(* CODESYS project cylinder.library
   DefaultNamespace: KOSTAL.AF2024.Drivers.Actuation.Cylinder
   DocFormat: reStructuredText
   Description: Handle a base cylinder device with two out and two input channels.
   Author: Frank Dümpelmann
   Title: KOSTAL.AF2024.Drivers.Actuation.Cylinder
   Version: 1.0.3.0
   Company: KOSTAL GmbH & Co.KG
   Placeholder: KOSTAL.AF2024.Drivers.Actuation.Cylinder

Project tree, tasks and I/O mapping:
  libraries: KOSTAL.AF2024.Core.functionResponse, 1.0.0.0 (KOSTAL GmbH & Co.KG); KOSTAL.AF2024.Core.ListOf, 1.0.0.0 (KOSTAL GmbH & Co.KG); KOSTAL.AF2024.Core.Process, 1.0.0.0 (KOSTAL GmbH & Co.KG); KOSTAL.AF2024.Core.Settings, 1.0.0.0 (KOSTAL GmbH & Co.KG); KOSTAL.AF2024.Core.Station, 1.0.0.0 (KOSTAL GmbH & Co.KG); KOSTAL.AF2024.Core.System, 1.0.0.0 (KOSTAL GmbH & Co.KG); KOSTAL.AF2024.Core.Text, 1.0.0.0 (KOSTAL GmbH & Co.KG); Tc2_Standard, 3.3.3.0 (Beckhoff Automation GmbH)
  Base/
    Cylinder_Base/
      function block _FB_Cylinder_Base [ST]: _fill, _mode, _moveTo_A, _moveTo_B, _pressureless, _set, conditionTime, conditionTime_ToA, conditionTime_ToB, NoLimitSwitch, sensor_A, sensor_B, valve_A, valve_B, FBmain
      interface _I_Cylinder_base: conditionTime, conditionTime_ToA, conditionTime_ToB, NoLimitSwitch, sensor_A, sensor_B, valve_A, valve_B, FBmain
      interface _I_Cylinder_base_RO: conditionTime, conditionTime_ToA, conditionTime_ToB, NoLimitSwitch, sensor_A, sensor_B, valve_A, valve_B
    Cylinder_Controlled_Base/
      function block _FB_Cylinder_Controlled_base [ST]: _manualMode_Set, _manualModeControl, _set, Error, Error_RO, errorText_overlap, errorText_timeout, ManualMode_Active, ManualMode_AutomaticRelease, ManualMode_Interlock, Name, Name_RO, overlapControl, timeout, timeoutControl, ManualMode_Reset, _fill, _moveTo_A, _moveTo_B, _pressureless, FBmain
      interface _I_Cylinder_Controlled_Base: ManualMode_Active, ManualMode_AutomaticRelease, ManualMode_Interlock, Error, Error_RO, errorText_overlap, errorText_timeout, Name, Name_RO, overlapControl, timeout, timeoutControl, ManualMode_Reset
      interface _I_Cylinder_Controlled_Base_RO: ManualMode_Active, ManualMode_AutomaticRelease, ManualMode_Interlock, Error_RO, errorText_overlap, errorText_timeout, Name_RO, overlapControl, timeout, timeoutControl
  DUT/
    Error/
      ListOf/
      interface I_T_Error: Clear, CopyFrom, active, text
      interface I_T_Error_CopyFrom: CopyFrom
      interface I_T_Error_RO: CopyTo, active, text
      function block T_Error [ST]: clear, CopyFrom, CopyTo, active, text
    Name/
      ListOf/
      interface I_T_Name: Clear, CopyFrom, device, sensor_A, sensor_B, valve_A, valve_B
      interface I_T_Name_CopyFrom: CopyFrom
      interface I_T_Name_RO: CopyTo, device, sensor_A, sensor_B, valve_A, valve_B
      function block T_Name [ST]: clear, CopyFrom, CopyTo, device, sensor_A, sensor_B, valve_A, valve_B
    StateMemory/
      ListOf/
        function block FB_ListOf_StateMemory [ST]: _get_I, _get_I_RO, _removePayLoad, _verifyMember, Add_DUT, Clear, CopyFrom, CopyTo, Delete_DUT, Find_DUT_byKey, Get_I, Get_I_RO, HasKey, Remove_DUT, MaxEntries, NumberOfMember
        interface I_ListOf_StateMemory: Add_DUT, Clear, CopyFrom, CopyTo, Delete_DUT, Get_I, Get_I_RO, NumberOfMember
        interface I_ListOf_StateMemory_CopyFrom: CopyFrom
        interface I_ListOf_StateMemory_RO: CopyTo, Get_I_RO, NumberOfMember
      interface I_T_StateMemory: Clear, CopyFrom, Key, Valve_A, Valve_B
      interface I_T_StateMemory_CopyFrom: CopyFrom
      interface I_T_StateMemory_RO: CopyTo, Key, Valve_A, Valve_B
      function block T_StateMemory [ST]: Clear, CopyFrom, CopyTo, Key, Valve_A, Valve_B
    TextHandler/
      function block FB_Text [ST]: AddVar, AddVar_UTF8, ClearVars, GetText
    data type _E_Mode
  POU/
    Cylinder/
      function block FB_Cylinder [ST]: Fill, moveTo_A, moveTo_B, Pressureless
      interface I_Cylinder: Fill, moveTo_A, moveTo_B, Pressureless
      interface I_Cylinder_RO
    Cylinder_Controlled/
      function block FB_Cylinder_Controlled [ST]: Fill, moveTo_A, moveTo_B, Pressureless
      interface I_Cylinder_Controlled: Fill, ManualMode_Reset, moveTo_A, moveTo_B, Pressureless
      interface I_Cylinder_Controlled_RO
    Cylinder_Step/
      function block FB_Cylinder_Step [ST]: FB_exit, FB_init, _addState, _StateHandling, _errorHandler, _execute, _mode, _parameterControl, ClearMemory, Fill, moveTo_A, moveTo_B, Pressureless, FBmain
      interface I_Cylinder_Step: Fill, moveTo_A, moveTo_B, Pressureless, ClearMemory
      data type ST_Manual
  Project Information/
    function F_GetCompany [ST]
    function F_GetTitle [ST]
    function F_GetVersion [ST]
  Version/
    global variables Global_Version
*)

// DUT/_E_Mode
(*
Description
===========
| Mode of cylinder control
| 0 = Normal: move to selected direction 
| 1 = Pressureless: close both valves
| 2 = Fill: open both valves  
*)
{attribute 'qualified_only'}
{attribute 'strict'}
TYPE _E_Mode :
	(
		NORMAL 			:= 0,
		PRESSURELESS	:= 1,
		FILL 			:= 2
	);
END_TYPE

// POU/Cylinder_Step/ST_Manual

TYPE ST_Manual :
STRUCT
	ManualValveMode 	: BOOL;
	ManualInterlock 	: BOOL;
	AutomaticRelease 	: BOOL;
	
	RequestManualOn		: BOOL;
	RequestManualOff	: BOOL;
	
	Valve_A				: BOOL;
	Valve_B				: BOOL;
	ResetCounter		: BYTE := 1;
	
END_STRUCT
END_TYPE

// Version/Global_Version
{attribute 'TcGenerated'}
{attribute 'no-analysis'}
{attribute 'linkalways'}
// This function has been automatically generated from the project information.
VAR_GLOBAL CONSTANT
	{attribute 'const_non_replaced'}
	stLibVersion_KOSTAL_AF2024_Drivers_Actuation_Cylinder : ST_LibVersion := (iMajor := 1, iMinor := 0, iBuild := 3, iRevision := 0, nFlags := 0, sVersion := '1.0.3.0');
END_VAR

// Base/Cylinder_Base/_FB_Cylinder_Base
{attribute 'enable_dynamic_creation'}
{attribute 'qualified_only'}
FUNCTION_BLOCK PUBLIC _FB_Cylinder_Base IMPLEMENTS _I_Cylinder_Base_RO, _I_Cylinder_Base

VAR CONSTANT
	_defTimeMin	: TIME:= TO_TIME(4294967295);	//T#0D0H0M0MS;	//define minimum default time
END_VAR

VAR
	_sensor_A	: BOOL;	//BOOL
	_sensor_B	: BOOL;	//BOOL
	_valve_A	: BOOL;	//BOOL
	_valve_B	: BOOL;	//BOOL

	_noLimitSwitch		: BOOL;
	
	_conditionTimer_moveToA	: TON;	//TON
	_conditionTime_ToA			: TIME	:= _defTimeMin;	//TIME	:= _defTimeMin - default = use common conditionTime

	_conditionTimer_moveToB	: TON;	//TON
	_conditionTime_ToB			: TIME	:= _defTimeMin;	//TIME	:= _defTimeMin - default = use common conditionTime

	_conditionTimer_moveProcess	: TON;	//TON
	_conditionTime							: TIME	:= T#100MS;	//TIME	:= T#100ms - default
	
END_VAR


METHOD PROTECTED _fill : BOOL

_fill:= FALSE;

_mode(_e_mode.FILL, FALSE, FALSE);

_conditionTimer_moveProcess.IN:= TRUE; 
_fill:= _conditionTimer_moveProcess.IN AND _conditionTimer_moveProcess.Q;
END_METHOD

METHOD PROTECTED _mode

VAR_INPUT
	mode	: _E_Mode;	//E_Mode
	to_A	: BOOL;	//BOOL
	to_B	: BOOL;	//BOOL
END_VAR
IF mode = _E_Mode.PRESSURELESS THEN

	_valve_A:= FALSE;
	_valve_B:= FALSE;

ELSIF mode = _E_Mode.FILL THEN

	_valve_A:= TRUE;
	_valve_B:= TRUE;

ELSE	//NORMAL

	_valve_A:= to_A;
	_valve_B:= to_B;
		
END_IF
END_METHOD


METHOD PROTECTED _moveTo_A : BOOL

_moveTo_A:= FALSE;

_mode(_E_Mode.NORMAL,TRUE, FALSE);

//_conditionTimer_moveToA.IN:= _sensor_A AND NOT (NOT _noSwitch AND _sensor_B);
_conditionTimer_moveToA.IN:= (_sensor_A AND NOT _sensor_B) OR _noLimitSwitch; 
 
_moveTo_A:= _conditionTimer_moveToA.IN AND _conditionTimer_moveToA.Q;
END_METHOD

METHOD PROTECTED _moveTo_B : BOOL

_moveTo_B:= FALSE;

_mode(_E_Mode.NORMAL, FALSE, TRUE);

_conditionTimer_moveToB.IN:= (_sensor_B AND NOT _sensor_A) OR _noLimitSwitch; 
_moveTo_B:= _conditionTimer_moveToB.IN AND _conditionTimer_moveToB.Q;
END_METHOD

METHOD PROTECTED _pressureless : BOOL

_pressureless:= FALSE;

_mode(_E_Mode.PRESSURELESS, FALSE, FALSE);

_conditionTimer_moveProcess.IN:= TRUE; 
_pressureless:= _conditionTimer_moveProcess.IN AND _conditionTimer_moveProcess.Q;
END_METHOD

METHOD PROTECTED _set
VAR_INPUT
END_VAR


IF _conditionTime_ToA = _defTimeMin THEN 	_conditionTimer_moveToA.PT:= _conditionTime;
ELSE																			_conditionTimer_moveToA.PT:= _conditionTime_ToA;
END_IF
_conditionTimer_moveToA();
_conditionTimer_moveToA.IN:= FALSE;	//default

IF _conditionTime_ToB = _defTimeMin THEN 	_conditionTimer_moveToB.PT:= _conditionTime;
ELSE																			_conditionTimer_moveToB.PT:= _conditionTime_ToB;
END_IF
_conditionTimer_moveToB();
_conditionTimer_moveToB.IN:= FALSE;	//default

_conditionTimer_moveProcess(IN:= , PT:= _conditionTime, Q=> , ET=> );
_conditionTimer_moveProcess.IN:= FALSE;	//default
END_METHOD

(*
Description
===========
| Minimum time before a movement function returns TRUE
*)
PROPERTY PUBLIC conditionTime : TIME
GET

conditionTime:= _conditionTime;
END_GET
SET

_conditionTime:= conditionTime;
END_SET
END_PROPERTY

(*
Description
===========
| Minimum time before a movement function returns TRUE
*)
PROPERTY PUBLIC conditionTime_ToA : TIME
GET

conditionTime_ToA:= _conditionTime_ToA;
END_GET
SET

_conditionTime_ToA:= conditionTime_ToA;
END_SET
END_PROPERTY

(*
Description
===========
| Minimum time before a movement function returns TRUE
*)
PROPERTY PUBLIC conditionTime_ToB : TIME
GET

conditionTime_ToB:= _conditionTime_ToB;
END_GET
SET

_conditionTime_ToB:= conditionTime_ToB;
END_SET
END_PROPERTY

(*
Description
===========
| TRUE: Both sensors active together result in a fault.
*)
PROPERTY PUBLIC NoLimitSwitch : BOOL
GET

NoLimitSwitch:= _noLimitSwitch;
END_GET
SET
_noLimitSwitch := NoLimitSwitch;
END_SET
END_PROPERTY

(*
Description
===========
| Sensor for home position
| Set TRUE if no sensor installed
*)
PROPERTY PUBLIC sensor_A : BOOL
GET

sensor_A:= _sensor_A;
END_GET
SET

_sensor_A:= sensor_A;
END_SET
END_PROPERTY

(*
Description
===========
| Sensor for work position
| Set TRUE if no sensor installed
*)
PROPERTY PUBLIC sensor_B : BOOL
GET

sensor_B:= _sensor_B;
END_GET
SET

_sensor_B:= sensor_B;
END_SET
END_PROPERTY

(*
Description
===========
| Valve to move cylinder to home position
*)
PROPERTY PUBLIC valve_A : BOOL
GET

valve_A:= _valve_A;
END_GET
SET

_valve_A:= valve_A;
END_SET
END_PROPERTY

(*
Description
===========
| Valve to move cylinder to work position
*)
PROPERTY PUBLIC valve_B : BOOL
GET

valve_B:= _valve_B;
END_GET
SET

_valve_B:= valve_B;
END_SET
END_PROPERTY

(*
Description
===========
| Main method, to be called cyclicly, e.g. in DeviceDefine
*)
METHOD PUBLIC FBmain
VAR_INPUT
END_VAR
	
_set();
END_METHOD

END_FUNCTION_BLOCK

// Base/Cylinder_Base/_I_Cylinder_base_RO
INTERFACE _I_Cylinder_base_RO EXTENDS KOSTAL_AF2024_Core_System.I_Interface

(*
Description
===========
| Minimum time before a movement function returns TRUE
*)
PROPERTY PUBLIC conditionTime : TIME
GET
END_GET
END_PROPERTY

(*
Description
===========
| Minimum time before a movement function returns TRUE
*)
PROPERTY PUBLIC conditionTime_ToA : TIME
GET
END_GET
END_PROPERTY

(*
Description
===========
| Minimum time before a movement function returns TRUE
*)
PROPERTY PUBLIC conditionTime_ToB : TIME
GET
END_GET
END_PROPERTY

(*
Description
===========
| TRUE: Both sensors active together result in a fault.
*)
PROPERTY PUBLIC NoLimitSwitch : BOOL
GET
END_GET
END_PROPERTY

(*
Description
===========
| Sensor for home position
| Set TRUE if no sensor installed
*)
PROPERTY PUBLIC sensor_A : BOOL
GET
END_GET
END_PROPERTY

(*
Description
===========
| Sensor for work position
| Set TRUE if no sensor installed
*)
PROPERTY PUBLIC sensor_B : BOOL
GET
END_GET
END_PROPERTY

(*
Description
===========
| Valve to move cylinder to home position
*)
PROPERTY PUBLIC valve_A : BOOL
GET
END_GET
END_PROPERTY

(*
Description
===========
| Valve to move cylinder to work position
*)
PROPERTY PUBLIC valve_B : BOOL
GET
END_GET
END_PROPERTY

END_INTERFACE

// Base/Cylinder_Base/_I_Cylinder_base
INTERFACE _I_Cylinder_base EXTENDS KOSTAL_AF2024_Core_System.I_Interface

(*
Description
===========
| Minimum time before a movement function returns TRUE
*)
PROPERTY PUBLIC conditionTime : TIME
GET
END_GET
SET
END_SET
END_PROPERTY

(*
Description
===========
| Minimum time before a movement function returns TRUE
*)
PROPERTY PUBLIC conditionTime_ToA : TIME
GET
END_GET
SET
END_SET
END_PROPERTY

(*
Description
===========
| Minimum time before a movement function returns TRUE
*)
PROPERTY PUBLIC conditionTime_ToB : TIME
GET
END_GET
SET
END_SET
END_PROPERTY

(*
Description
===========
| TRUE: Ignore Sensor inputs.
*)
PROPERTY PUBLIC NoLimitSwitch : BOOL
GET
END_GET
SET
END_SET
END_PROPERTY

(*
Description
===========
| Sensor for home position
| Set TRUE if no sensor installed
*)
PROPERTY PUBLIC sensor_A : BOOL
GET
END_GET
SET
END_SET
END_PROPERTY

(*
Description
===========
| Sensor for work position
| Set TRUE if no sensor installed
*)
PROPERTY PUBLIC sensor_B : BOOL
GET
END_GET
SET
END_SET
END_PROPERTY

(*
Description
===========
| Valve to move cylinder to home position
*)
PROPERTY PUBLIC valve_A : BOOL
GET
END_GET
SET
END_SET
END_PROPERTY

(*
Description
===========
| Valve to move cylinder to work position
*)
PROPERTY PUBLIC valve_B : BOOL
GET
END_GET
SET
END_SET
END_PROPERTY

(*
Description
===========
| Main method, to be called cyclicly, e.g. in DeviceDefine
*)
METHOD PUBLIC FBmain
VAR_INPUT
END_VAR
END_METHOD

END_INTERFACE

// Base/Cylinder_Controlled_Base/_FB_Cylinder_Controlled_base
{attribute 'enable_dynamic_creation'}
{attribute 'qualified_only'}
FUNCTION_BLOCK ABSTRACT _FB_Cylinder_Controlled_base EXTENDS _FB_Cylinder_Base IMPLEMENTS _I_Cylinder_Controlled_Base_RO, _I_Cylinder_Controlled_Base
VAR_INPUT
END_VAR
VAR_OUTPUT
END_VAR
VAR
	_timeOut			: TIME	:= T#5S;	//- default
	_timeOutTimer	: TON;
	
	_timeoutControl	: BOOL;
	_overlapControl	: BOOL;
	
	_errorText_timeout	: WSTRING;
	_errorText_overlap	: WSTRING;

	_Name		:	T_Name;
	_error	: T_Error;
	
	_textHandler	:FB_Text;
	
	//Manual control from HMI
	_automatic_A			: BOOL;
	_automatic_B			: BOOL;
	{attribute 'Cylinder_2024_V1'}
	_manual	: ST_Manual;
	
END_VAR

(*
Description
===========
| (De)activate manual valve mode
| Parameters:
| 	state : bool : TRUE = activate, FALSE = deactivate
*)
METHOD protected _manualMode_Set
VAR_INPUT
	state : bool;
END_VAR
//IF state THEN
//	_automatic_A := _valve_A;	//Store valve states before going to manual
//	_automatic_B := _valve_B;
////	_manual.ManualValveMode := TRUE;
////ELSE
////	_automatic_A 		:= FALSE;
////	_automatic_B 		:= FALSE;
////	_manual.ManualValveMode 	:= FALSE;
//END_IF
_manual.ManualValveMode := state;
END_METHOD

METHOD PROTECTED _manualModeControl
VAR_INPUT
END_VAR
IF NOT _manual.ManualValveMode THEN //Store valve states if not in manual
	_automatic_A := _valve_A;	
	_automatic_B := _valve_B;
END_IF

_manual.AutomaticRelease := (NOT (_valve_A XOR _automatic_A) AND NOT (_valve_B XOR _automatic_B));

IF _manual.RequestManualOn AND NOT _manual.ManualInterlock AND NOT _manual.ManualValveMode THEN
	//_manualMode_Set(TRUE);
	_manual.Valve_A := _valve_A;
	_manual.Valve_B := _valve_B;
	_manual.ManualValveMode := TRUE;
ELSIF _manual.RequestManualOff AND _manual.AutomaticRelease AND _manual.ManualValveMode THEN
//	_manualMode_Set(FALSE);
	_manual.ManualValveMode := FALSE;
END_IF

IF _manual.ManualValveMode AND NOT _manual.ManualInterlock THEN
	_valve_A := _manual.Valve_A;
	_valve_B := _manual.Valve_B;
END_IF
END_METHOD

METHOD PROTECTED _set
VAR_INPUT
END_VAR


SUPER^._set();


_timeOutTimer(PT:= _timeOut);
_error.active:= _timeOutTimer.Q;

_timeOutTimer.IN:= FALSE;	//default

_error.clear();
END_METHOD

(*
Description
===========
| See documentation of FB_error
| **Attention:** Errors are reset in FB_Main. Check errors before FB_Main is called!
*)
PROPERTY PUBLIC Error : I_T_Error
GET

Error := _error;
END_GET
END_PROPERTY

PROPERTY PUBLIC Error_RO : I_T_Error_RO
GET

Error_RO:= _error;
END_GET
END_PROPERTY

(*
Description
===========
| Message Text for overlap error
*)
PROPERTY PUBLIC errorText_overlap : KOSTAL_AF2024_Core_Settings.T_MaxString
GET

errorText_overlap:= _errorText_overlap;
END_GET
SET

_errorText_overlap:= errorText_overlap;
END_SET
END_PROPERTY

(*
Description
===========
| Message Text for timeout error
*)
PROPERTY PUBLIC errorText_timeout : KOSTAL_AF2024_Core_Settings.T_MaxString
GET

errorText_Timeout:= _errorText_timeout;
END_GET
SET

_errorText_Timeout:= errorText_timeout;
END_SET
END_PROPERTY

(*
Description
===========
| TRUE if manual control is activated for this cylinder
*)
PROPERTY PUBLIC ManualMode_Active : BOOL
GET
ManualMode_Active := _manual.ManualValveMode;
END_GET
END_PROPERTY

(*
Description
===========
| True if manual valve state equals automatic valve state
| -> Enable automatic mode 
*)
// 
PROPERTY PUBLIC ManualMode_AutomaticRelease : BOOL
GET
ManualMode_AutomaticRelease := _manual.AutomaticRelease;
END_GET
END_PROPERTY

(*
Description
===========
| Interlock manual cylinder control
*)
PROPERTY PUBLIC ManualMode_Interlock : BOOL
GET
ManualMode_Interlock := _manual.ManualInterlock;
END_GET
SET
_manual.ManualInterlock := ManualMode_Interlock;
END_SET
END_PROPERTY

PROPERTY PUBLIC Name : I_T_Name
GET

Name:= _Name;
END_GET
END_PROPERTY

(*
Description
===========
| Naming of cilinders and componets (see documentation of FB_name)
*)
PROPERTY PUBLIC Name_RO : I_T_Name_RO
GET

Name_RO := _Name;
END_GET
END_PROPERTY

(*
Description
===========
| TRUE: Both sensors active together result in a fault.
*)
PROPERTY PUBLIC overlapControl : BOOL
GET

overlapControl:= _overlapControl;
END_GET
SET

_overlapControl:= overlapControl;
END_SET
END_PROPERTY

(*
Description
===========
| Time for timeoutControl
| Default: 5s
*)
PROPERTY PUBLIC timeout : TIME
GET

timeout:= _timeOut;
END_GET
SET

_timeout:= timeOut;
END_SET
END_PROPERTY

(*
Description
===========
| TRUE: generate error when movement is not finished after a certain time
*)
PROPERTY PUBLIC timeoutControl : BOOL
GET

timeoutControl:= _timeoutControl;
END_GET
SET

_timeoutControl:= timeoutControl;
END_SET
END_PROPERTY

METHOD Public ManualMode_Reset : BOOL
VAR_INPUT
END_VAR

_manualMode_Set(FALSE);
_manual.Valve_A := _manual.Valve_B := FALSE;
_manual.ResetCounter := LIMIT(1, _manual.ResetCounter + 1, 254);

ManualMode_Reset := THIS^._pressureless();
END_METHOD

METHOD PROTECTED _fill : BOOL

_fill:= SUPER^._fill();

_timeOutTimer(IN:= NOT _conditionTimer_moveProcess.IN AND _timeoutControl, PT:= _timeOut);

IF _overlapControl AND _sensor_A AND _sensor_B AND NOT _noLimitSwitch THEN

	_error.active:= TRUE;

	_textHandler.clearVars();
	_textHandler.AddVar(Name_RO.sensor_A);
	_textHandler.AddVar(Name_RO.sensor_B);
	_error.text:=  _textHandler.getText(errorText_overlap);

ELSE

	_error.active:= FALSE;
	_error.text:= "";
	
END_IF
END_METHOD

METHOD PROTECTED _moveTo_A : BOOL

_moveTo_A:= SUPER^._moveTo_A();


_timeOutTimer(IN:= NOT _conditionTimer_moveToA.IN AND _timeoutControl, PT:= _timeOut);

IF _overlapControl AND _sensor_A AND _sensor_B AND NOT _noLimitSwitch THEN

	_error.active:= TRUE;
	
	_textHandler.clearVars();
	_textHandler.AddVar(Name_RO.sensor_A);
	_textHandler.AddVar(Name_RO.sensor_B);
	_error.text:=  _textHandler.GetText(errorText_overlap);

ELSIF _timeOutTimer.Q THEN

	_error.active:= TRUE;

	_textHandler.clearVars();
	_textHandler.AddVar(Name_RO.sensor_A);
	_error.text:=  _textHandler.GetText(errorText_timeout);

ELSE

	_error.active:= FALSE;
	_error.text:= "";
	
END_IF
END_METHOD

METHOD PROTECTED _moveTo_B : BOOL

_moveTo_B:= SUPER^._moveTo_B();


_timeOutTimer(IN:= NOT _conditionTimer_moveToB.IN AND _timeoutControl, PT:= _timeOut);

IF _overlapControl AND _sensor_A AND _sensor_B AND NOT _noLimitSwitch THEN

	_error.active:= TRUE;

	_textHandler.clearVars();
	_textHandler.AddVar(Name_RO.sensor_A);
	_textHandler.AddVar(Name_RO.sensor_B);
	_error.text:=  _textHandler.getText(errorText_overlap);

ELSIF _timeOutTimer.Q THEN

	_error.active:= TRUE;

	_textHandler.clearVars();
	_textHandler.AddVar(Name_RO.sensor_B);
	_error.text:=  _textHandler.getText(errorText_timeout);

ELSE

	_error.active:= FALSE;
	_error.text:= "";
	
END_IF
END_METHOD

METHOD PROTECTED _pressureless : BOOL

_pressureless:= SUPER^._pressureless();

_timeOutTimer(IN:= NOT _conditionTimer_moveProcess.IN AND _timeoutControl, PT:= _timeOut);

IF _overlapControl AND _sensor_A AND _sensor_B AND NOT _noLimitSwitch THEN

	_error.active:= TRUE;

	_textHandler.clearVars();
	_textHandler.AddVar(Name_RO.sensor_A);
	_textHandler.AddVar(Name_RO.sensor_B);
	_error.text:=  _textHandler.getText(errorText_overlap);

ELSE

	_error.active:= FALSE;
	_error.text:= "";
	
END_IF
END_METHOD

(*
Description
===========
| Main method, to be called cyclicly, e.g. in DeviceDefine
*)
METHOD PUBLIC FBmain
VAR_INPUT
END_VAR
SUPER^.FBmain();
_manualModeControl();
END_METHOD

END_FUNCTION_BLOCK

// Base/Cylinder_Controlled_Base/_I_Cylinder_Controlled_Base_RO
INTERFACE _I_Cylinder_Controlled_Base_RO EXTENDS _I_Cylinder_Base_RO

PROPERTY PUBLIC ManualMode_Active : BOOL
GET
END_GET
END_PROPERTY

//Manual valve state = automatic valve state -> Release automatic mode
PROPERTY PUBLIC ManualMode_AutomaticRelease : BOOL
GET
END_GET
END_PROPERTY

PROPERTY PUBLIC ManualMode_Interlock : BOOL
GET
END_GET
END_PROPERTY

PROPERTY PUBLIC Error_RO : I_T_Error_RO
GET
END_GET
END_PROPERTY

(*
Description
===========
| Message Text for overlap error
*)
PROPERTY PUBLIC errorText_overlap : KOSTAL_AF2024_Core_Settings.T_MaxString
GET
END_GET
SET
END_SET
END_PROPERTY

(*
Description
===========
| Message Text for timeout error
*)
PROPERTY PUBLIC errorText_timeout : KOSTAL_AF2024_Core_Settings.T_MaxString
GET
END_GET
END_PROPERTY

(*
Description
===========
| Naming of cilinders and componets (see documentation of FB_name)
*)
{attribute 'obsolete' := 'use instead property IName or method LinkName()!'} 
PROPERTY PUBLIC Name_RO : I_T_Name_RO
GET
END_GET
END_PROPERTY

(*
Description
===========
| TRUE: Both sensors active together result in a fault.
*)
PROPERTY PUBLIC overlapControl : BOOL
GET
END_GET
END_PROPERTY

(*
Description
===========
| Time for timeoutControl
| Default: 5s
*)
PROPERTY PUBLIC timeout : TIME
GET
END_GET
END_PROPERTY

(*
Description
===========
| TRUE: generate error when movement is not finished after a certain time
*)
PROPERTY PUBLIC timeoutControl : BOOL
GET
END_GET
END_PROPERTY

END_INTERFACE

// DUT/Error/I_T_Error_RO
(*
	Read only Interface from DUT
*)
INTERFACE I_T_Error_RO  EXTENDS KOSTAL_AF2024_Core_System.I_Interface

METHOD PUBLIC CopyTo
VAR_INPUT
	IN	: I_T_Error_CopyFrom;
END_VAR
END_METHOD

(*
Description
===========
| Error is active
*)
PROPERTY PUBLIC active : BOOL
GET
END_GET
END_PROPERTY

(*
Description
===========
| Text of error message
*)
PROPERTY PUBLIC text : KOSTAL_AF2024_Core_Settings.T_MaxString
GET
END_GET
END_PROPERTY

END_INTERFACE

// DUT/Error/I_T_Error_CopyFrom
INTERFACE I_T_Error_CopyFrom EXTENDS KOSTAL_AF2024_Core_System.I_Interface

METHOD PUBLIC CopyFrom
VAR_INPUT
	IN	: I_T_Error_RO;
END_VAR
END_METHOD

END_INTERFACE

// DUT/Name/I_T_Name_RO
(*
	Read only Interface from DUT
*)
INTERFACE I_T_Name_RO  EXTENDS KOSTAL_AF2024_Core_System.I_Interface

METHOD PUBLIC CopyTo
VAR_INPUT
	IN	: I_T_Name_CopyFrom;
END_VAR
END_METHOD

(*
Description
===========
| Name of the cylinder
*)
PROPERTY PUBLIC device : KOSTAL_AF2024_Core_Settings.T_MaxString
GET
END_GET
END_PROPERTY

(*
Description
===========
| Name of the cylinder's home position sensor
*)
PROPERTY PUBLIC sensor_A : KOSTAL_AF2024_Core_Settings.T_MaxString
GET
END_GET
END_PROPERTY

(*
Description
===========
| Name of the cylinder's work position sensor
*)
PROPERTY PUBLIC sensor_B : KOSTAL_AF2024_Core_Settings.T_MaxString
GET
END_GET
END_PROPERTY

(*
Description
===========
| Name of the cylinder's home position actuator
*)
PROPERTY PUBLIC valve_A : KOSTAL_AF2024_Core_Settings.T_MaxString
GET
END_GET
END_PROPERTY

(*
Description
===========
| Name of the cylinder's work position actuator
*)
PROPERTY PUBLIC valve_B : KOSTAL_AF2024_Core_Settings.T_MaxString
GET
END_GET
END_PROPERTY

END_INTERFACE

// DUT/Name/I_T_Name_CopyFrom
INTERFACE I_T_Name_CopyFrom EXTENDS KOSTAL_AF2024_Core_System.I_Interface

METHOD PUBLIC CopyFrom
VAR_INPUT
	IN	: I_T_Name_RO;
END_VAR
END_METHOD

END_INTERFACE

// Base/Cylinder_Controlled_Base/_I_Cylinder_Controlled_Base
INTERFACE _I_Cylinder_Controlled_Base EXTENDS _I_Cylinder_base

PROPERTY PUBLIC ManualMode_Active : BOOL
GET
END_GET
END_PROPERTY

//Manual valve state = automatic valve state -> Release automatic mode
PROPERTY PUBLIC ManualMode_AutomaticRelease : BOOL
GET
END_GET
END_PROPERTY

PROPERTY PUBLIC ManualMode_Interlock : BOOL
GET
END_GET
SET
END_SET
END_PROPERTY

(*
Description
===========
| See documentation of FB_error
| **Attention:** Errors are reset in FB_Main. Check errors before FB_Main is called!
*)
PROPERTY PUBLIC Error : I_T_Error
GET
END_GET
END_PROPERTY

PROPERTY PUBLIC Error_RO : I_T_Error_RO
GET
END_GET
END_PROPERTY

(*
Description
===========
| Message Text for overlap error
*)
PROPERTY PUBLIC errorText_overlap : KOSTAL_AF2024_Core_Settings.T_MaxString
GET
END_GET
SET
END_SET
END_PROPERTY

(*
Description
===========
| Message Text for timeout error
*)
PROPERTY PUBLIC errorText_timeout : KOSTAL_AF2024_Core_Settings.T_MaxString
GET
END_GET
SET
END_SET
END_PROPERTY

PROPERTY PUBLIC Name : I_T_Name
GET
END_GET
END_PROPERTY

(*
Description
===========
| Naming of cilinders and componets (see documentation of FB_name)
*)
{attribute 'obsolete' := 'use instead property IName or method LinkName()!'} 
PROPERTY PUBLIC Name_RO : I_T_Name_RO
GET
END_GET
END_PROPERTY

(*
Description
===========
| TRUE: Both sensors active together result in a fault.
*)
PROPERTY PUBLIC overlapControl : BOOL
GET
END_GET
SET
END_SET
END_PROPERTY

(*
Description
===========
| Time for timeoutControl
| Default: 5s
*)
PROPERTY PUBLIC timeout : TIME
GET
END_GET
SET
END_SET
END_PROPERTY

(*
Description
===========
| TRUE: generate error when movement is not finished after a certain time
*)
PROPERTY PUBLIC timeoutControl : BOOL
GET
END_GET
SET
END_SET
END_PROPERTY

METHOD Public ManualMode_Reset : BOOL
VAR_INPUT
END_VAR
END_METHOD

END_INTERFACE

// DUT/Error/I_T_Error
(*
	Full qualified access Interface from DUT
*)
INTERFACE I_T_Error EXTENDS I_T_Error_RO

METHOD PUBLIC Clear
END_METHOD

METHOD PUBLIC CopyFrom
VAR_INPUT
	IN	: I_T_Error_RO;
END_VAR
END_METHOD

(*
Description
===========
| Error is active
*)
PROPERTY PUBLIC active : BOOL
SET
END_SET
END_PROPERTY

(*
Description
===========
| Text of error message
*)
PROPERTY PUBLIC text : KOSTAL_AF2024_Core_Settings.T_MaxString
SET
END_SET
END_PROPERTY

END_INTERFACE

// DUT/Name/I_T_Name
(*
	Full qualified access Interface from DUT
*)
INTERFACE I_T_Name EXTENDS I_T_Name_RO

METHOD PUBLIC Clear : BOOL
VAR_INPUT
END_VAR
END_METHOD

METHOD PUBLIC CopyFrom
VAR_INPUT
	IN	: I_T_Name_RO;
END_VAR
END_METHOD

(*
Description
===========
| Name of the cylinder
*)
PROPERTY PUBLIC device : KOSTAL_AF2024_Core_Settings.T_MaxString
SET
END_SET
END_PROPERTY

(*
Description
===========
| Name of the cylinder's home position sensor
*)
PROPERTY PUBLIC sensor_A : KOSTAL_AF2024_Core_Settings.T_MaxString
SET
END_SET
END_PROPERTY

(*
Description
===========
| Name of the cylinder's work position sensor
*)
PROPERTY PUBLIC sensor_B : KOSTAL_AF2024_Core_Settings.T_MaxString
SET
END_SET
END_PROPERTY

(*
Description
===========
| Name of the cylinder's home position actuator
*)
PROPERTY PUBLIC valve_A : KOSTAL_AF2024_Core_Settings.T_MaxString
SET
END_SET
END_PROPERTY

(*
Description
===========
| Name of the cylinder's work position actuator
*)
PROPERTY PUBLIC valve_B : KOSTAL_AF2024_Core_Settings.T_MaxString
SET
END_SET
END_PROPERTY

END_INTERFACE

// DUT/Name/T_Name
(*

:Author: Frank Dümpelmann <f.duempelmann@kostal.com>, Martin Hundt <m.hundt@kostal.com>
:Date: 2018-11-19

Function
========
| Data type for naming cylinders and their components (valves, sensors)

Methods and Properties
======================
| See bottom of this document for a detailed description of each method or property
*)

{attribute 'enable_dynamic_creation'}
{attribute 'qualified_only'}
FUNCTION_BLOCK T_Name IMPLEMENTS I_T_Name_RO, I_T_Name, I_T_Name_CopyFrom

VAR
	_device		: KOSTAL_AF2024_Core_Settings.T_MaxString;
	_sensor_A	: KOSTAL_AF2024_Core_Settings.T_MaxString;
	_sensor_B	: KOSTAL_AF2024_Core_Settings.T_MaxString;
	_valve_A	: KOSTAL_AF2024_Core_Settings.T_MaxString;
	_valve_B	: KOSTAL_AF2024_Core_Settings.T_MaxString;
END_VAR

(*
Description
===========
| Clear all naming
*)
METHOD clear : BOOL
VAR_INPUT
END_VAR

_device		:= "";
_sensor_A	:= "";
_sensor_B	:= "";
_valve_A	:= "";
_valve_B	:= "";
END_METHOD

METHOD PUBLIC CopyFrom
VAR_INPUT
	IN	: I_T_Name_RO;
END_VAR

IF IN = 0 THEN RETURN;	END_IF

_device		:= IN.device;
_sensor_A	:= IN.sensor_A;
_sensor_B	:= IN.sensor_B;
_valve_A	:= IN.valve_A;
_valve_B	:= IN.valve_B;
END_METHOD

METHOD PUBLIC CopyTo
VAR_INPUT
	IN	: I_T_Name_CopyFrom;
END_VAR

IF IN = 0 THEN RETURN;	END_IF

IN.CopyFrom(THIS^);
END_METHOD

(*
Description
===========
| Name of the cylinder
*)
PROPERTY PUBLIC device : KOSTAL_AF2024_Core_Settings.T_MaxString
GET

device:= _device;
END_GET
SET

_device:= device;
END_SET
END_PROPERTY

(*
Description
===========
| Name of the cylinder's home position sensor
*)
PROPERTY PUBLIC sensor_A : KOSTAL_AF2024_Core_Settings.T_MaxString
GET

sensor_A:= _sensor_A;
END_GET
SET

_sensor_A:= sensor_A;
END_SET
END_PROPERTY

(*
Description
===========
| Name of the cylinder's work position sensor
*)
PROPERTY PUBLIC sensor_B : KOSTAL_AF2024_Core_Settings.T_MaxString
GET

sensor_B:= _sensor_B;
END_GET
SET

_sensor_B:= sensor_B;
END_SET
END_PROPERTY

(*
Description
===========
| Name of the cylinder's home position actuator
*)
PROPERTY PUBLIC valve_A : KOSTAL_AF2024_Core_Settings.T_MaxString
GET

valve_A:= _valve_A;
END_GET
SET

_valve_A:= valve_A;
END_SET
END_PROPERTY

(*
Description
===========
| Name of the cylinder's work position actuator
*)
PROPERTY PUBLIC valve_B : KOSTAL_AF2024_Core_Settings.T_MaxString
GET

valve_B:= _valve_B;
END_GET
SET

_valve_B:= valve_B;
END_SET
END_PROPERTY

END_FUNCTION_BLOCK

// DUT/Error/T_Error
(*

:Author: Frank Dümpelmann <f.duempelmann@kostal.com>, Martin Hundt <m.hundt@kostal.com>
:Date: 2018-11-19

Function
========
| Data type for error messages

Methods and Properties
======================
| See bottom of this document for a detailed description of each method or property
*)
{attribute 'enable_dynamic_creation'}
{attribute 'qualified_only'}
FUNCTION_BLOCK T_Error IMPLEMENTS I_T_Error_RO, I_T_Error, I_T_Error_CopyFrom

VAR
	_active	: BOOL;
	_text		: KOSTAL_AF2024_Core_Settings.T_MaxString;
END_VAR

METHOD PUBLIC Clear

_active	:= FALSE;
_text		:= "";
END_METHOD

METHOD PUBLIC CopyFrom
VAR_INPUT
	IN	: I_T_Error_RO;
END_VAR

IF IN = 0 THEN RETURN;	END_IF

_active	:= IN.active;
_text		:= IN.text;
END_METHOD

METHOD PUBLIC CopyTo
VAR_INPUT
	IN	: I_T_Error_CopyFrom;
END_VAR

IF IN = 0 THEN RETURN;	END_IF

IN.CopyFrom(THIS^);
END_METHOD

(*
Description
===========
| Error is active
*)
PROPERTY PUBLIC active : BOOL
GET

active:= _active;
END_GET
SET

_active:= active;
END_SET
END_PROPERTY

(*
Description
===========
| Text of error message
*)
PROPERTY PUBLIC text : KOSTAL_AF2024_Core_Settings.T_MaxString
GET

text:= _text;
END_GET
SET

_text:= text;
END_SET
END_PROPERTY

END_FUNCTION_BLOCK

// DUT/TextHandler/FB_Text
FUNCTION_BLOCK INTERNAL FB_Text EXTENDS Kostal_AF2024_Core_Text._FB_Base
VAR_INPUT
END_VAR
VAR_OUTPUT
END_VAR
VAR
END_VAR

METHOD AddVar : BOOL
VAR_INPUT
	Text	: KOSTAL_AF2024_Core_Settings.T_MaxString;
END_VAR

AddVar:= _Variables.addLine(Text);
END_METHOD

METHOD AddVar_UTF8 : BOOL
VAR_INPUT
	Text	: KOSTAL_AF2024_Core_Settings.T_MaxString;
END_VAR



AddVar_UTF8:= _Variables.addLine(Text);
END_METHOD

METHOD ClearVars

_Variables.clear();
END_METHOD

METHOD GetText : KOSTAL_AF2024_Core_Settings.T_MaxString

VAR_INPUT
	Text	: KOSTAL_AF2024_Core_Settings.T_MaxString;
END_VAR

GetText:= "";

IF Text = "" THEN RETURN;	END_IF

GetText:= _combine(Text);
END_METHOD

END_FUNCTION_BLOCK

// DUT/StateMemory/ListOf/FB_ListOf_StateMemory
(*
	A template for creating a list of typed classes (FBs)
*)
FUNCTION_BLOCK FB_ListOf_StateMemory EXTENDS KOSTAL_AF2024_Core_ListOf._FB_Object_Base  IMPLEMENTS I_ListOf_StateMemory_RO, I_ListOf_StateMemory_CopyFrom, I_ListOf_StateMemory

VAR
	//Use the {_Dummy} to ensure that a valid interface is always returned.
	_Dummy			: T_StateMemory;
	_MaxEntries	: UDINT:= UDINT#128;
END_VAR

(*
	Returns the typed owner interface in the reference variable.
	In the event of an error, the return value becomes FALSE and the interface refers to the {_Dummy}.
*)
METHOD PROTECTED _get_I : BOOL

VAR_INPUT
	Member		: KOSTAL_AF2024_Core_System.I_Interface;
	rFound_I	: REFERENCE TO I_T_StateMemory;
	rResult		: KOSTAL_AF2024_Core_functionResponse.I_T_functionResponse_Owner;
END_VAR

VAR
	_iObj			: I_T_StateMemory;
	_Success	: BOOL;
END_VAR

IF NOT SUPER^._verifyMember(Member, rResult)	THEN 
	IF __ISVALIDREF(rFound_I)	THEN	rFound_I:= _Dummy;	END_IF
	RETURN;	
END_IF

_Success:= __QUERYINTERFACE(Member, _iObj);

//return dummy if no valid DUT is found
IF NOT _Success OR (_iObj = 0)	THEN	

	IF __ISVALIDREF(rFound_I)	THEN	rFound_I:= _Dummy;	END_IF	
	IF rResult <> 0						THEN	rResult.success:= FALSE;	
																	rResult.status:= "__QueryInterface failed - return Dummy";	
	END_IF	

	RETURN;	

END_IF

IF __ISVALIDREF(rFound_I)	THEN	rFound_I:= _iObj;	END_IF
IF rResult <> 0						THEN	rResult.success:= TRUE;
																rResult.status:= "Successful";
END_IF

_get_I:= TRUE;
END_METHOD

(*
	Returns the typed interface in the reference variable.
	In the event of an error, the return value becomes FALSE and the interface refers to the {_Dummy}.
*)
METHOD PROTECTED _get_I_RO : BOOL

VAR_INPUT
	Member		: KOSTAL_AF2024_Core_System.I_Interface;
	rFound_I	: REFERENCE TO I_T_StateMemory_RO;
	rResult		: KOSTAL_AF2024_Core_functionResponse.I_T_functionResponse_Owner;
END_VAR

VAR
	_iObj	: I_T_StateMemory_RO;
	_Success: BOOL;
END_VAR

IF NOT SUPER^._verifyMember(Member, rResult)	THEN 
	IF __ISVALIDREF(rFound_I)	THEN	rFound_I:= _Dummy;	END_IF
	RETURN;	
END_IF

_Success:= __QUERYINTERFACE(Member, _iObj);

//return dummy if no valid DUT is found
IF NOT _Success OR (_iObj = 0)	THEN	

	IF __ISVALIDREF(rFound_I)	THEN	rFound_I:= _Dummy;	END_IF	
	IF rResult <> 0						THEN	rResult.success:= FALSE;		
																	rResult.status:= "__QueryInterface failed - return Dummy";	
	END_IF	

	RETURN;	

END_IF

IF __ISVALIDREF(rFound_I)	THEN	rFound_I:= _iObj;	END_IF
IF rResult <> 0						THEN	rResult.success:= TRUE;
																rResult.status:= "Successful";
END_IF

_get_I_RO:= TRUE;
END_METHOD

(*
	Cleans the custom class {FB_DUT} and removes it from memory.
*)
METHOD PROTECTED  _removePayLoad : BOOL
VAR_INPUT
	Member	: KOSTAL_AF2024_Core_System.I_Interface;
	Result	: KOSTAL_AF2024_Core_functionResponse.I_T_functionResponse_Owner;
END_VAR

VAR
	_iObj			: I_T_StateMemory;
	_pFB_DUT	:	POINTER TO T_StateMemory;
	_Success	: BOOL;
END_VAR


IF NOT SUPER^._removePayload(Member, Result)	THEN RETURN;	END_IF

_Success:= __QUERYINTERFACE(Member, _iObj);

IF NOT _Success	THEN	RETURN;	END_IF
IF _iObj = 0		THEN	RETURN;	END_IF

_iObj.Clear();

_Success  := __QUERYPOINTER(_iObj, _pFB_DUT);

IF NOT _Success	THEN	RETURN;	END_IF
IF _pFB_DUT = 0	THEN	RETURN;	END_IF

__DELETE(_pFB_DUT);
END_METHOD

(*
	Overload the method from the base class to verify the custom interface. 
	The local method {_get_I_Owner()} is used for this.
*)
METHOD PROTECTED _verifyMember : BOOL
VAR_INPUT
	Member	: KOSTAL_AF2024_Core_System.I_Interface;
	Result	: KOSTAL_AF2024_Core_functionResponse.I_T_functionResponse_Owner;
END_VAR


_verifyMember:= _get_I(Member, 0, Result);
END_METHOD

(*
	Add a new instance of FB_Dut and copy content from [IN] to the new instance
*)
METHOD PUBLIC Add_DUT : BOOL
VAR_INPUT
	IN				: I_T_StateMemory_RO;
	Response	: KOSTAL_AF2024_Core_functionResponse.I_T_functionResponse_Owner;
END_VAR

VAR
	_iDUT	: I_T_StateMemory;
	_pDUT: POINTER TO T_StateMemory;
	_response: KOSTAL_AF2024_Core_functionResponse.T_functionResponse;
	_udi: UDINT;
END_VAR

_response.clear();

IF IN = 0 THEN
	IF Response <> 0 THEN	Response.success:= FALSE;	Response.status:= "IN Parameter is invalid";	END_IF
	RETURN;
END_IF

IF _Count	> _MaxEntries THEN 
	IF Response <> 0 THEN	Response.success:= FALSE;	Response.status:= "Max entries overflow";	END_IF
	RETURN;	
END_IF

_pDUT:= __NEW(T_StateMemory);

IF _pDUT = 0 THEN
	_response.status:= "cannot create new object";
	IF Response <> 0 THEN	Response.CopyFrom(_response);	END_IF
	RETURN;
END_IF

_pDUT^.CopyFrom(IN);

SUPER^._addMember(_pDUT^, _response);

IF Response <> 0 THEN	Response.CopyFrom(_response);	END_IF

Add_DUT:= _response.success;
END_METHOD

(*
	Makes the protected method public.
*)
METHOD Clear

SUPER^._clear();
END_METHOD

(*
	Copies the contents of another list {IN} into its own memory.
*)
METHOD PUBLIC CopyFrom
VAR_INPUT
	IN	: I_ListOf_StateMemory_RO;
END_VAR

VAR
	_udi	: UDINT;
	_IDUT	: I_T_StateMemory_RO;
END_VAR
IF IN = 0 THEN RETURN;	END_IF

_clear();

FOR _udi:= 1 TO IN.NumberOfMember DO
	IF IN.Get_I_RO(_udi, _IDUT, 0)	THEN	Add_DUT(_IDUT, 0);	END_IF
END_FOR
END_METHOD

(*
	Copies the own content into another list created at the parameter {IN}.
*)
METHOD PUBLIC CopyTo
VAR_INPUT
	IN	: I_ListOf_StateMemory_CopyFrom;
END_VAR

IF IN = 0 THEN RETURN;	END_IF

IN.CopyFrom(THIS^);
END_METHOD

(*
	Deletes the class specified with the {Number} from the list.
*)
METHOD PUBLIC Delete_DUT : BOOL
VAR_INPUT
	Number		: UDINT;	//Number of DUT in List
	Response	: KOSTAL_AF2024_Core_functionResponse.I_T_functionResponse_Owner;
END_VAR

VAR
	_response	: KOSTAL_AF2024_Core_functionResponse.T_functionResponse;
	_Success	: BOOL;
	_Member		: KOSTAL_AF2024_Core_System.I_Interface;
END_VAR

IF Number = 0 THEN
	_response.clear(); _response.status:= "Number is out of range (1..n)"; 
	IF Response <> 0 THEN	Response.CopyFrom(_response);	END_IF
	RETURN;
END_IF

Delete_DUT:= SUPER^._removeMemberByIndex(Number - 1, _response);

IF Response <> 0 THEN	Response.CopyFrom(_response);	END_IF

Delete_DUT:= _response.success;
END_METHOD

METHOD Find_DUT_byKey : BOOL
VAR_INPUT
	Key	: ULINT;
	rFound_I	: REFERENCE TO I_T_StateMemory_RO;
END_VAR

VAR
	_udi: UDINT;
	_iMem				: KOSTAL_AF2024_Core_System.I_Interface;
	_iStateMem	: I_T_StateMemory_RO;
	_Success: BOOL;
END_VAR

IF _Count = 0 THEN	rFound_I:= _Dummy;	Find_DUT_byKey:= FALSE;	RETURN;	END_IF

FOR _udi:= _Count - 1 TO 0 BY -1 DO 

	IF _findMemberByIndex(_udi, _iMem, 0) AND_THEN _iMem <> 0 THEN 

		_Success:= __QUERYINTERFACE(_iMem, _iStateMem);
		
		//return dummy if no valid DUT is found
		IF NOT _Success OR_ELSE (_iStateMem = 0)	THEN	
		
			IF __ISVALIDREF(rFound_I)	THEN	rFound_I:= _Dummy;	Find_DUT_byKey:= FALSE; END_IF	
			RETURN;	

		ELSE

			IF _iStateMem.Key = Key THEN
					
				IF __ISVALIDREF(rFound_I) THEN	rFound_I:= _iStateMem;	Find_DUT_byKey:= TRUE;	RETURN;	END_IF
		
			END_IF


		END_IF
	
	ELSE

		IF __ISVALIDREF(rFound_I)	THEN	rFound_I:= _Dummy;	Find_DUT_byKey:= FALSE; END_IF	
		RETURN;	
	
	END_IF
	
END_FOR

IF __ISVALIDREF(rFound_I) THEN	rFound_I:= _Dummy;	Find_DUT_byKey:= FALSE;	RETURN;	END_IF
END_METHOD

(*
	Get full access to content of Member with {Number}
*) 
METHOD Get_I : BOOL

VAR_INPUT
	Number		: UDINT;
	rFound_I	: REFERENCE TO I_T_StateMemory;
	Response	: KOSTAL_AF2024_Core_functionResponse.I_T_functionResponse_Owner;
END_VAR

VAR
	_Member				: KOSTAL_AF2024_Core_System.I_Interface;
	_response			: KOSTAL_AF2024_Core_functionResponse.T_functionResponse;
END_VAR

IF Number = 0 THEN
	_response.clear(); _response.status:= "Number is out of range (1..n)"; 
	IF Response <> 0 THEN	Response.CopyFrom(_response);	END_IF
	RETURN;
END_IF

IF NOT SUPER^._findMemberByIndex(Number - 1, _Member, Response) THEN

 IF __ISVALIDREF(rFound_I) THEN	rFound_I:= _Dummy;	END_IF

ELSE

	Get_I:= _get_I(_Member, rFound_I, Response);
	
END_IF
END_METHOD

(*
	Get readonly access to content of Member with {Number}
*) 
METHOD Get_I_RO : BOOL

VAR_INPUT
	Number		: UDINT;
	rFound_I	: REFERENCE TO I_T_StateMemory_RO;
	Response	: KOSTAL_AF2024_Core_functionResponse.I_T_functionResponse_Owner;
END_VAR

VAR
	_Member		: KOSTAL_AF2024_Core_System.I_Interface;
	_response	: KOSTAL_AF2024_Core_functionResponse.T_functionResponse;
END_VAR
IF Number = 0 THEN
	_response.clear(); _response.status:= "Number is out of range (1..n)"; 
	IF Response <> 0 THEN	Response.CopyFrom(_response);	END_IF
	RETURN;
END_IF

IF NOT SUPER^._findMemberByIndex(Number - 1, _Member, Response) THEN

 IF __ISVALIDREF(rFound_I) THEN	rFound_I:= _Dummy;	END_IF

ELSE

	Get_I_RO:= _get_I_RO(_Member, rFound_I, Response);
	
END_IF
END_METHOD

METHOD PUBLIC HasKey : BOOL
VAR_INPUT
	IN	: ULINT;
END_VAR


VAR
	_udi: UDINT;
	_Mem: I_T_StateMemory;
END_VAR

FOR _udi:= 1 TO _Count DO
	IF Get_I(_udi, _Mem, 0) (*AND_THEN (_Mem <> 0)*) AND_THEN _Mem.Key = IN THEN HasKey:= TRUE; RETURN; END_IF
END_FOR

HasKey:= FALSE;
END_METHOD

(*
	Deletes the class specified with the {Number} from the list.
*)
METHOD PUBLIC Remove_DUT : BOOL
VAR_INPUT
	Member		: I_T_StateMemory_RO;
	Response	: KOSTAL_AF2024_Core_functionResponse.I_T_functionResponse_Owner;
END_VAR

VAR
	_response	: KOSTAL_AF2024_Core_functionResponse.T_functionResponse;
	_Success	: BOOL;
	_Member		: KOSTAL_AF2024_Core_System.I_Interface;
END_VAR

IF Member = 0 THEN
	_response.clear(); _response.status:= "Parameter Member is invalid"; 
	IF Response <> 0 THEN	Response.CopyFrom(_response);	END_IF
	RETURN;
END_IF

Remove_DUT:= SUPER^._removeMember(Member, _response);

IF Response <> 0 THEN	Response.CopyFrom(_response);	END_IF

Remove_DUT:= _response.success;
END_METHOD

PROPERTY PUBLIC MaxEntries : UDINT
GET

MaxEntries:= _MaxEntries;
END_GET
SET

_MaxEntries:= MaxEntries;
END_SET
END_PROPERTY

(*
	Number of Member in list.
*)
PROPERTY NumberOfMember : UDINT
GET

NumberOfMember:= SUPER^._NumberOfMember;
END_GET
END_PROPERTY

END_FUNCTION_BLOCK

// DUT/StateMemory/ListOf/I_ListOf_StateMemory_RO
(*
	Read only Interface from List of DUT
*)
INTERFACE I_ListOf_StateMemory_RO EXTENDS KOSTAL_AF2024_Core_ListOf._I_Object_Base

METHOD PUBLIC CopyTo
VAR_INPUT
	IN	: I_ListOf_StateMemory_CopyFrom;
END_VAR
END_METHOD

METHOD Get_I_RO : BOOL

VAR_INPUT
	Number		: UDINT;
	rFound_I	: REFERENCE TO I_T_StateMemory_RO;
	Response	: KOSTAL_AF2024_Core_functionResponse.I_T_functionResponse_Owner;
END_VAR
END_METHOD

PROPERTY NumberOfMember : UDINT
GET
END_GET
END_PROPERTY

END_INTERFACE

// DUT/StateMemory/ListOf/I_ListOf_StateMemory_CopyFrom
(*
	The class implementing this interface can take over the contents from another instance with the same interface {I_DUT}.
	Typing takes place in the method.
*)
INTERFACE I_ListOf_StateMemory_CopyFrom EXTENDS KOSTAL_AF2024_Core_System.I_Interface

(*
	Copies the contents of another list {IN} into its own memory.
*)
METHOD PUBLIC CopyFrom
VAR_INPUT
	IN	: I_ListOf_StateMemory_RO;
END_VAR
END_METHOD

END_INTERFACE

// DUT/StateMemory/I_T_StateMemory_RO
INTERFACE I_T_StateMemory_RO EXTENDS KOSTAL_AF2024_Core_System.I_Interface

METHOD PUBLIC CopyTo : BOOL
VAR_INPUT
	IN	: I_T_StateMemory_CopyFrom;
END_VAR
END_METHOD

PROPERTY PUBLIC Key : ULINT
GET
END_GET
END_PROPERTY

PROPERTY PUBLIC Valve_A : BOOL
GET
END_GET
END_PROPERTY

PROPERTY PUBLIC Valve_B : BOOL
GET
END_GET
END_PROPERTY

END_INTERFACE

// DUT/StateMemory/I_T_StateMemory_CopyFrom
INTERFACE I_T_StateMemory_CopyFrom EXTENDS KOSTAL_AF2024_Core_System.I_Interface

METHOD PUBLIC CopyFrom	:	BOOL
VAR_INPUT
	IN	: I_T_StateMemory_RO;
END_VAR
END_METHOD

END_INTERFACE

// DUT/StateMemory/ListOf/I_ListOf_StateMemory
(*
	Full qualified access Interface from List of DUT
*)
INTERFACE I_ListOf_StateMemory EXTENDS KOSTAL_AF2024_Core_ListOf._I_Object_Base_Owner

//Add a new instance of FB_Dut and copy content from [IN] to the new instance
METHOD PUBLIC Add_DUT : BOOL
VAR_INPUT
	IN				: I_T_StateMemory_RO;
	Response	: KOSTAL_AF2024_Core_functionResponse.I_T_functionResponse_Owner;
END_VAR
END_METHOD

METHOD Clear
VAR_INPUT
END_VAR
END_METHOD

METHOD PUBLIC CopyFrom
VAR_INPUT
	IN	: I_ListOf_StateMemory_RO;
END_VAR
END_METHOD

METHOD PUBLIC CopyTo
VAR_INPUT
	IN	: I_ListOf_StateMemory_CopyFrom;
END_VAR
END_METHOD

METHOD PUBLIC Delete_DUT : BOOL
VAR_INPUT
	Number	: UDINT;	//Number of DUT in List
	Response	: KOSTAL_AF2024_Core_functionResponse.I_T_functionResponse_Owner;
END_VAR
END_METHOD

//Get full access to content 
METHOD Get_I : BOOL

VAR_INPUT
	Number		: UDINT;
	rFound_I	: REFERENCE TO I_T_StateMemory;
	Response	: KOSTAL_AF2024_Core_functionResponse.I_T_functionResponse_Owner;
END_VAR
END_METHOD

METHOD Get_I_RO : BOOL

VAR_INPUT
	Number		: UDINT;
	rFound_I	: REFERENCE TO I_T_StateMemory_RO;
	Response	: KOSTAL_AF2024_Core_functionResponse.I_T_functionResponse_Owner;
END_VAR
END_METHOD

PROPERTY NumberOfMember : UDINT
GET
END_GET
END_PROPERTY

END_INTERFACE

// DUT/StateMemory/I_T_StateMemory
INTERFACE I_T_StateMemory EXTENDS I_T_StateMemory_RO

METHOD PUBLIC Clear
END_METHOD

METHOD PUBLIC CopyFrom	:	BOOL
VAR_INPUT
	IN	: I_T_StateMemory_RO;
END_VAR
END_METHOD

PROPERTY PUBLIC Key : ULINT
SET
END_SET
END_PROPERTY

PROPERTY PUBLIC Valve_A : BOOL
SET
END_SET
END_PROPERTY

PROPERTY PUBLIC Valve_B : BOOL
SET
END_SET
END_PROPERTY

END_INTERFACE

// DUT/StateMemory/T_StateMemory
{attribute 'enable_dynamic_creation'}
FUNCTION_BLOCK PUBLIC T_StateMemory IMPLEMENTS I_T_StateMemory_RO, I_T_StateMemory, I_T_StateMemory_CopyFrom
VAR
	_Key			: ULINT;	//Contains the unique step key
	_Valve_A	: BOOL;		//State of valve "A" when stepping into the execution
	_Valve_B	: BOOL;		//State of valve "B" when stepping into the execution
END_VAR

METHOD PUBLIC Clear

_Key			:= ULINT#0;
_Valve_A	:= FALSE;
_Valve_B	:= FALSE;
END_METHOD

METHOD PUBLIC CopyFrom	:	BOOL
VAR_INPUT
	IN	: I_T_StateMemory_RO;
END_VAR

IF IN = 0 THEN RETURN;	END_IF

_Key			:= IN.Key;
_Valve_A	:= IN.Valve_A;
_Valve_B	:= IN.Valve_B;

CopyFrom:= TRUE;
END_METHOD

METHOD PUBLIC CopyTo : BOOL
VAR_INPUT
	IN	: I_T_StateMemory_CopyFrom;
END_VAR

IF IN = 0 THEN RETURN;	END_IF

IN.CopyFrom(THIS^);

CopyTo:= TRUE;
END_METHOD

PROPERTY PUBLIC Key : ULINT
GET

Key:= _Key;
END_GET
SET

_Key:= Key;
END_SET
END_PROPERTY

PROPERTY PUBLIC Valve_A : BOOL
GET

Valve_A:= _Valve_A;
END_GET
SET

_Valve_A:= Valve_A;
END_SET
END_PROPERTY

PROPERTY PUBLIC Valve_B : BOOL
GET

Valve_B:= _Valve_B;
END_GET
SET

_Valve_B:= Valve_B;
END_SET
END_PROPERTY

END_FUNCTION_BLOCK

// POU/Cylinder/FB_Cylinder
(*

:Author: Frank Dümpelmann <f.duempelmann@kostal.com>, Martin Hundt <m.hundt@kostal.com>
:Date: 2018-11-19

Function
========
| Function block representing basic functions of a cylinder with max. two valves and two sensors

Usage notes
===============
| Asyncronous function block: FBmain() method must be called cyclicly
| Call function moveTo_A to go to home position
| Call function moveTo_B to go to work position
| Call function moveProcess to set the modes pressureless, fill or freeze

Methods and Properties
======================
| See bottom of this document for a detailed description of each method or property
| Methods starting with an underline(_) are internally used and can be ignored by the user


*)
{attribute 'enable_dynamic_creation'}
{attribute 'qualified_only'}
FUNCTION_BLOCK PUBLIC FB_Cylinder EXTENDS _FB_Cylinder_Base IMPLEMENTS I_Cylinder_RO, I_Cylinder

VAR
	
END_VAR

(*
Description
===========
| Fill the Cylinder (both valves open)

| Returns: BOOL - Function carried out successfully
*)
METHOD PUBLIC Fill : BOOL

fill:=SUPER^._fill();
END_METHOD

(*
Description
===========
| Move cylinder to home position
| Returns: BOOL - Move carried out successfully
*)
METHOD PUBLIC moveTo_A : BOOL

moveTo_A:= SUPER^._moveTo_A();
END_METHOD

(*
Description
===========
| Move cylinder to work position
| Returns: BOOL - Move carried out successfully
*)
METHOD PUBLIC moveTo_B : BOOL
moveTo_B:= SUPER^._moveTo_B();
END_METHOD

(*
Description
===========
| Set the Cylinder Pressureless (both valves closed)

| Returns: BOOL - Function carried out successfully
*)
METHOD PUBLIC Pressureless : BOOL

pressureless:=SUPER^._pressureless();
END_METHOD

END_FUNCTION_BLOCK

// POU/Cylinder/I_Cylinder_RO
INTERFACE I_Cylinder_RO EXTENDS _I_Cylinder_base_RO

END_INTERFACE

// POU/Cylinder/I_Cylinder
INTERFACE I_Cylinder EXTENDS _I_Cylinder_base

(*
Description
===========
| Fill the Cylinder (both valves open)

| Returns: BOOL - Function carried out successfully
*)
METHOD PUBLIC Fill : BOOL
END_METHOD

(*
Description
===========
| Move cylinder to home position
| Returns: BOOL - Move carried out successfully
*)
METHOD PUBLIC moveTo_A : BOOL
END_METHOD

(*
Description
===========
| Move cylinder to work position
| Returns: BOOL - Move carried out successfully
*)
METHOD PUBLIC moveTo_B : BOOL
END_METHOD

(*
Description
===========
| Set the Cylinder Pressureless (both valves closed)

| Returns: BOOL - Function carried out successfully
*)
METHOD PUBLIC Pressureless : BOOL
END_METHOD

END_INTERFACE

// POU/Cylinder_Controlled/FB_Cylinder_Controlled
(*

:Author: Frank Dümpelmann <f.duempelmann@kostal.com>, Martin Hundt <m.hundt@kostal.com>
:Date: 2018-11-19

Function
========
| Extends FB_Cylinder with functions for timeout control, naming and error messaging
| See also documentation of FB_Cylinder

Usage notes
===============
| Asyncronous function block: FBmain() method must be called cyclicly
| Call function moveTo_A to go to home position
| Call function moveTo_B to go to work position
| Call function moveProcess to set the modes pressureless, fill or freeze
| **Attention:** Errors are reset in FBmain. Check errors before FBmain is called!

Methods and Properties
======================
| See bottom of this document for a detailed description of each method or property
| Methods starting with an underline(_) are internally used and can be ignored by the user

*)
{attribute 'enable_dynamic_creation'}
{attribute 'qualified_only'}
FUNCTION_BLOCK PUBLIC FB_Cylinder_Controlled EXTENDS _FB_Cylinder_Controlled_base IMPLEMENTS I_Cylinder_Controlled_RO, I_Cylinder_Controlled
VAR_INPUT
END_VAR
VAR_OUTPUT
END_VAR
VAR
	
	
END_VAR

(*
Description
===========
| Fill the Cylinder (both valves open)

| Returns: BOOL - Function carried out successfully
*)
METHOD PUBLIC Fill : BOOL

fill:=SUPER^._fill();
END_METHOD

(*
Description
===========
| Move cylinder to home position
| Returns: BOOL - Move carried out successfully
*)
METHOD PUBLIC moveTo_A : BOOL

moveTo_A:= SUPER^._moveTo_A();
END_METHOD

(*
Description
===========
| Move cylinder to work position
| Returns: BOOL - Move carried out successfully
*)
METHOD PUBLIC moveTo_B : BOOL
moveTo_B:= SUPER^._moveTo_B();
END_METHOD

(*
Description
===========
| Set the Cylinder Pressureless (both valves closed)

| Returns: BOOL - Function carried out successfully
*)
METHOD PUBLIC Pressureless : BOOL

pressureless:=SUPER^._pressureless();
END_METHOD

END_FUNCTION_BLOCK

// POU/Cylinder_Controlled/I_Cylinder_Controlled_RO
INTERFACE I_Cylinder_Controlled_RO EXTENDS _I_Cylinder_Controlled_Base_RO

END_INTERFACE

// POU/Cylinder_Controlled/I_Cylinder_Controlled
INTERFACE I_Cylinder_Controlled EXTENDS _I_Cylinder_Controlled_Base

(*
Description
===========
| Fill the Cylinder (both valves open)

| Returns: BOOL - Function carried out successfully
*)
METHOD PUBLIC Fill : BOOL
END_METHOD

METHOD PUBLIC ManualMode_Reset : BOOL
VAR_INPUT
END_VAR
END_METHOD

(*
Description
===========
| Move cylinder to home position
| Returns: BOOL - Move carried out successfully
*)
METHOD PUBLIC moveTo_A : BOOL
END_METHOD

(*
Description
===========
| Move cylinder to work position
| Returns: BOOL - Move carried out successfully
*)
METHOD PUBLIC moveTo_B : BOOL
END_METHOD

(*
Description
===========
| Set the Cylinder Pressureless (both valves closed)

| Returns: BOOL - Function carried out successfully
*)
METHOD PUBLIC Pressureless : BOOL
END_METHOD

END_INTERFACE

// POU/Cylinder_Step/FB_Cylinder_Step
{attribute 'qualified_only'}
FUNCTION_BLOCK PUBLIC FB_Cylinder_Step EXTENDS _FB_Cylinder_Controlled_base IMPLEMENTS I_Cylinder_Step

VAR
	_Station				: KOSTAL_AF2024_Core_Station.I_Station_Controlled_Owner;
	_StateMemory			: FB_ListOf_StateMemory;

	_execution				:	BOOL;

	_stepMemoryCountOld		: UDINT;

END_VAR

METHOD FB_exit : BOOL
VAR_INPUT
	bInCopyCode : BOOL; // if TRUE, the exit method is called for exiting an instance that is copied afterwards (online change).
END_VAR

_StateMemory.Clear();
END_METHOD

METHOD FB_init : BOOL
VAR_INPUT
	bInitRetains : BOOL; // if TRUE, the retain variables are initialized (warm start / cold start)
	bInCopyCode : BOOL;  // if TRUE, the instance afterwards gets moved into the copy code (online change)
	station	: KOSTAL_AF2024_Core_Station.I_Station_Controlled_Owner;
END_VAR
_Station := station;
_StateMemory.Clear();
END_METHOD

METHOD PROTECTED _addState : BOOL

VAR
	_Mem		: 	KOSTAL_AF2024_Core_Process.I_T_StepMemory_RO;
	_Cstate	:	T_StateMemory;
	_resp		: KOSTAL_AF2024_Core_functionResponse.T_functionResponse;
END_VAR

//if thie step key does not exist in list of state memory then ...	
IF _Station.Step.StepMemory_RO.Get_I_RO(_Station.Step.StepMemory_RO.NumberOfMember, _Mem, 0) 
AND_THEN NOT _StateMemory.HasKey(_Mem.RegKey)
THEN

	//try to create a stateMemory item with the key from toplevel stepMemory	
	_Cstate.Key		:= _Mem.RegKey;
	_Cstate.Valve_A	:= _valve_A;
	_Cstate.Valve_B	:= _valve_B;

	IF NOT _StateMemory.Add_DUT(_Cstate, _resp)	THEN	

		_Station.Message_Owner.clear();
		_Station.Message_Owner.line_01:= _Name.device;
		_Station.Message_Owner.line_02:= _resp.status;
		IF NOT _Station.Condition.isError() THEN	
			_Station.LogText(_Station.Message.toString());	
		END_IF
		_Station.Condition_Owner.setMessage(_Station.Condition.PriorityLevel_Error, _Station.Message);
		_station.Step_Owner.StepMemory.Clear();
		_StateMemory.Clear();

	END_IF

END_IF
END_METHOD

//Call up this method to update the step memory.
METHOD PROTECTED _StateHandling

VAR
	_StepMem	: KOSTAL_AF2024_Core_Process.I_T_StepMemory_RO;
	_Mem			: T_StateMemory;
	_IMem			: I_T_StateMemory_RO;
	_resp			: KOSTAL_AF2024_Core_functionResponse.T_functionResponse;
END_VAR


IF _Station.Step.BackwardDone THEN

	IF _StateMemory.Find_DUT_byKey(_Station.Step.LastUsedKey, _IMem) AND_THEN _IMem <> 0 THEN

		_valve_A:= _IMem.Valve_A;
		_valve_B:= _IMem.Valve_B;
		
		_StateMemory.Remove_DUT(_IMem, 0);
		
	ELSE
			
		_Station.Message_Owner.clear();
		_Station.Message_Owner.line_01:= _Name.device;
		_Station.Message_Owner.line_02:= "no StateMemory Element abvailable";
		IF NOT _Station.Condition.isError() THEN	
			_Station.LogText(_Station.Message.toString());	
		END_IF
		_Station.Condition_Owner.setMessage(_Station.Condition.PriorityLevel_Error, _Station.Message);

	END_IF

END_IF
END_METHOD

METHOD PROTECTED _errorHandler
VAR_INPUT
END_VAR


IF _error.active THEN

	_Station.Message_Owner.clear();
	_Station.Message_Owner.line_01:= _error.text;

	IF NOT _Station.Condition.isError() THEN	_Station.LogText(_Station.Message.toString());	END_IF 
	
	_Station.Condition_Owner.setMessage(_Station.Condition_Owner.PriorityLevel_Error, _Station.Message);
	
END_IF
END_METHOD

METHOD PROTECTED _execute : BOOL

IF NOT _parameterControl()	THEN RETURN; END_IF
IF _execution				THEN RETURN; END_IF

IF _Station.Step.toggle 		THEN	
	_addState();	
END_IF

_execution:= TRUE;
END_METHOD

METHOD PROTECTED _mode
VAR_INPUT
	mode	: _E_Mode;	//E_Mode
	to_A	: BOOL;	//BOOL
	to_B	: BOOL;	//BOOL
END_VAR
IF _manual.ManualValveMode THEN //Ignore moveTo... commands in manual state  
	;
ELSE
	SUPER^._mode(mode, to_A, to_B);
END_IF
END_METHOD

(*
| returns TRUE if parameter are valid
*)
METHOD PROTECTED _parameterControl : BOOL

_parameterControl:= (_Station <> 0);
END_METHOD

//Call up this method to delete the saved status history.
METHOD PUBLIC ClearMemory

_StateMemory.Clear();
END_METHOD

(*
Description
===========
| Fill the Cylinder (both valves open)
| Parameters:
|		jumpAddress	: INT - Address of next Step. 0 = +1
| 		stepRelease : BOOL - TRUE = Go to next step after process is finished
| Returns: BOOL - Function carried out successfully
*)
METHOD PUBLIC Fill : BOOL

VAR_INPUT
	jumpAddress	: INT;		
	stepRelease	: BOOL;		
END_VAR
IF NOT _parameterControl() THEN	RETURN; END_IF

_execute();

Fill:= SUPER^._fill();

_errorHandler();

IF NOT stepRelease THEN	_StateHandling();	RETURN;	END_IF

_Station.Step_Owner.Condition		:= Fill;
_Station.Step_Owner.JumpAddress	:= jumpAddress;

_Station.Step_Owner.Control();

_StateHandling();
END_METHOD

(*
Description
===========
| Move cylinder to home position
| Parameters:
|		jumpAddress	: INT - Address of next Step. 0 = +1
| 		stepRelease : BOOL - TRUE = Go to next step after process is finished
| Returns: BOOL - Move carried out successfully
*)
METHOD PUBLIC moveTo_A : BOOL
VAR_INPUT
	jumpAddress	: INT;		
	stepRelease	: BOOL;		
END_VAR
IF NOT _parameterControl() THEN	RETURN; END_IF

_execute();

moveTo_A:= SUPER^._moveTo_A();

_errorHandler();

IF NOT stepRelease THEN	
	_StateHandling();	
	RETURN;	
END_IF

_Station.Step_Owner.Condition		:= moveTo_A;
_Station.Step_Owner.JumpAddress	:= jumpAddress;

_Station.Step_Owner.Control();

_StateHandling();
END_METHOD

(*
Description
===========
| Move cylinder to work position
| Parameters:
|		jumpAddress	: INT - Address of next Step. 0 = +1
| 		stepRelease : BOOL - TRUE = Go to next step after process is finished
| Returns: BOOL - Move carried out successfully
*)
METHOD PUBLIC moveTo_B : BOOL
VAR_INPUT
	jumpAddress	: INT;		
	stepRelease	: BOOL;		
END_VAR
IF NOT _parameterControl() THEN	RETURN; END_IF

_execute();

moveTo_B:= SUPER^._moveTo_B();

_errorHandler();

IF NOT stepRelease THEN	_StateHandling();	RETURN;	END_IF

_Station.Step_Owner.Condition		:= moveTo_B;
_Station.Step_Owner.JumpAddress	:= jumpAddress;

_Station.Step_Owner.Control();

_StateHandling();
END_METHOD

(*
Description
===========
| Set the Cylinder Pressureless (both valves closed)
| Parameters:
|		jumpAddress	: INT - Address of next Step. 0 = +1
| 		stepRelease : BOOL - TRUE = Go to next step after process is finished
| Returns: BOOL - Function carried out successfully
*)
METHOD PUBLIC Pressureless : BOOL

VAR_INPUT
	jumpAddress	: INT;		
	stepRelease	: BOOL;		
END_VAR
IF NOT _parameterControl() THEN	RETURN; END_IF

_execute();

Pressureless:= SUPER^._pressureless();

_errorHandler();

IF NOT stepRelease THEN	_StateHandling();	RETURN;	END_IF

_Station.Step_Owner.Condition		:= Pressureless;
_Station.Step_Owner.JumpAddress	:= jumpAddress;

_Station.Step_Owner.Control();

_StateHandling();
END_METHOD

(*
Description
===========
| Main method, to be called cyclicly, e.g. in DeviceDefine
*)
METHOD PUBLIC FBmain
VAR_INPUT
END_VAR

SUPER^.FBmain();

//_manualModeControl();

_execution:= FALSE;

IF NOT _parameterControl() THEN	RETURN; END_IF

IF _StateMemory.NumberOfMember > 0 AND_THEN _Station.Step.StepMemory_RO.NumberOfMember < _stepMemoryCountOld THEN 
	_StateMemory.Clear();	
END_IF

_stepMemoryCountOld := _Station.Step.StepMemory_RO.NumberOfMember;
END_METHOD

END_FUNCTION_BLOCK

// POU/Cylinder_Step/I_Cylinder_Step
INTERFACE I_Cylinder_Step EXTENDS _I_Cylinder_Controlled_Base

(*
Description
===========
| Fill the Cylinder (both valves open)
| Parameters:
|		jumpAddress	: INT - Address of next Step. 0 = +1
| 		stepRelease : BOOL - TRUE = Go to next step after process is finished
| Returns: BOOL - Function carried out successfully
*)
METHOD PUBLIC Fill : BOOL

VAR_INPUT
	jumpAddress	: INT;		
	stepRelease	: BOOL;		
END_VAR
END_METHOD

(*
Description
===========
| Move cylinder to home position
| Parameters:
|		jumpAddress	: INT - Address of next Step. 0 = +1
| 		stepRelease : BOOL - TRUE = Go to next step after process is finished
| Returns: BOOL - Move carried out successfully
*)
METHOD PUBLIC moveTo_A : BOOL
VAR_INPUT
	jumpAddress	: INT;		
	stepRelease	: BOOL;		
END_VAR
END_METHOD

(*
Description
===========
| Move cylinder to work position
| Parameters:
|		jumpAddress	: INT - Address of next Step. 0 = +1
| 		stepRelease : BOOL - TRUE = Go to next step after process is finished
| Returns: BOOL - Move carried out successfully
*)
METHOD PUBLIC moveTo_B : BOOL
VAR_INPUT
	jumpAddress	: INT;		
	stepRelease	: BOOL;		
END_VAR
END_METHOD

(*
Description
===========
| Set the Cylinder Pressureless (both valves closed)
| Parameters:
|		jumpAddress	: INT - Address of next Step. 0 = +1
| 		stepRelease : BOOL - TRUE = Go to next step after process is finished
| Returns: BOOL - Function carried out successfully
*)
METHOD PUBLIC Pressureless : BOOL

VAR_INPUT
	jumpAddress	: INT;		
	stepRelease	: BOOL;		
END_VAR
END_METHOD

//Call up this method to delete the saved status history.
METHOD PUBLIC ClearMemory
END_METHOD

END_INTERFACE

// Project Information/F_GetCompany
// This function has been automatically generated from the project information.
{attribute 'signature_flag' := '1073741824'}
{attribute 'TcGenerated'}
{attribute 'no-analysis'}
FUNCTION F_GetCompany : WSTRING
VAR_INPUT
	
END_VAR

F_GetCompany := "KOSTAL GmbH & Co.KG";

END_FUNCTION

// Project Information/F_GetTitle
// This function has been automatically generated from the project information.
{attribute 'signature_flag' := '1073741824'}
{attribute 'TcGenerated'}
{attribute 'no-analysis'}
FUNCTION F_GetTitle : WSTRING
VAR_INPUT
	
END_VAR

F_GetTitle := "KOSTAL.AF2024.Drivers.Actuation.Cylinder";

END_FUNCTION

// Project Information/F_GetVersion
// This function has been automatically generated from the project information.
{attribute 'signature_flag' := '1073741824'}
{attribute 'TcGenerated'}
{attribute 'no-analysis'}
FUNCTION F_GetVersion : ST_LibVersion
VAR_INPUT
	
END_VAR

F_GetVersion.iMajor := 1;
F_GetVersion.iMinor := 0;
F_GetVersion.iBuild := 3;
F_GetVersion.iRevision := 0;
F_GetVersion.sVersion := '1.0.3.0';
F_GetVersion.nFlags := 0;

END_FUNCTION
